(* IEC 61131-3 sources: kns-port-domestic/targets/astra/src/POUs/Station/FB_PumpRotation, 14 files *)

(* ---- FB_PumpRotation.decl.st ---- *)
// Назначение: роли насосов, чередование и ограничение непрерывной работы (04 §5, §8). Запросы
//             получают насосы с ролями Lead и Assist; роли работающих по запросу насосов
//             сохраняются; недостающая роль — сначала ReadyToStart, затем доступные в паузе,
//             внутри группы — по eRotation (RunHours, Cyclic, Fixed); в ПИД ведущим — насос со
//             связью с ПЧ. Новый запрос — не раньше tStagger после предыдущего (если тот ещё
//             запрошен). Снятие роли: RunHours — насос с большей наработкой, Cyclic/Fixed —
//             подпорный. Отказавший насос теряет запрос сразу. Передача роли с перекрытием
//             tOverlap после tMaxContRun (событие 101007), повтор через STN_HANDOVER_RETRY.
//             uiRequestLimit (последовательный пуск) ограничивает новые запросы: насосы, уже
//             работающие по запросу (подхват при старте ПЛК), им не снимаются.
// Автор:      kr0nsch
// Версия:     0.1.0
// Документ:   docs/DESIGN.md, раздел 6.5; docs/04_algorithms.md, разделы 5, 8
FUNCTION_BLOCK FB_PumpRotation
VAR_INPUT
    xEnable          : BOOL;        // станция в «Автомате» (иначе запросов нет, роли считаются)
    uiRequired       : UINT;        // от действующего управления, 0…STN_PUMP_COUNT
    uiRequestLimit   : UINT;        // FB_PowerRestore: сколько запросов можно выдать
    xRequireComm     : BOOL;        // eControlAct = LevelPid: ведущий — только со связью
    xHandoverAllowed : BOOL;        // не Emergency, Float, Restart
    xAdopt           : BOOL;        // импульс: роли получают работающие насосы (вход в «Автомат», смена управления)
    axAdoptRun       : ARRAY[1..GVL_Const.STN_PUMP_COUNT] OF BOOL;  // «работает» для xAdopt (старт: GVL_IO.xP10n_RFB)
    aitfPump         : ARRAY[1..GVL_Const.STN_PUMP_COUNT] OF PL.I_MotorVfd;
    axCommOk         : ARRAY[1..GVL_Const.STN_PUMP_COUNT] OF BOOL;
    itfTime          : PL.I_TimeSource;
    itfEvents        : I_StationEventSink;
END_VAR
VAR_IN_OUT CONSTANT
    stCfg : ST_StationCfg;          // eRotation, uiDutyMax, tMaxContRun, tOverlap, tStagger
END_VAR
VAR_IN_OUT
    stRetain : ST_StationRetain;    // uiNextLead (Cyclic)
END_VAR
VAR_OUTPUT
    axRun              : ARRAY[1..GVL_Const.STN_PUMP_COUNT] OF BOOL;   // → fbP10n.xAutoRun
    aeRole             : ARRAY[1..GVL_Const.STN_PUMP_COUNT] OF E_PumpRole;
    uiLead             : UINT;
    uiAvailable        : UINT;      // Available
    uiRunning          : UINT;      // Running в любом режиме
    uiForeign          : UINT;      // работают не в Auto (сторонние, 04 §5.1)
    uiRequests         : UINT;      // запросы: не больше MAX(0, uiRequired - uiForeign), новые — до uiRequestLimit
    uiRunningRequested : UINT;      // запрошены и работают по ОС (для FB_PowerRestore)
    xHandover          : BOOL;      // идёт передача роли (перекрытие)
    xStaggerWait       : BOOL;      // новый запрос ждёт tStagger
END_VAR
VAR
    // снимок насосов этого вызова (методы читают его, а не интерфейсы)
    axAvail       : ARRAY[1..GVL_Const.STN_PUMP_COUNT] OF BOOL;    // Available
    axRunning     : ARRAY[1..GVL_Const.STN_PUMP_COUNT] OF BOOL;    // Running
    axReady       : ARRAY[1..GVL_Const.STN_PUMP_COUNT] OF BOOL;    // ReadyToStart
    audiHours     : ARRAY[1..GVL_Const.STN_PUMP_COUNT] OF UDINT;   // RunSeconds
    audiStarts    : ARRAY[1..GVL_Const.STN_PUMP_COUNT] OF UDINT;   // Starts
    audiCurRun    : ARRAY[1..GVL_Const.STN_PUMP_COUNT] OF UDINT;   // CurrentRunSeconds
    axForeign     : ARRAY[1..GVL_Const.STN_PUMP_COUNT] OF BOOL;    // работает не в Auto
    // запросы и роли
    axReq         : ARRAY[1..GVL_Const.STN_PUMP_COUNT] OF BOOL;    // запрос (роль Lead или Assist)
    audiReqSeq    : ARRAY[1..GVL_Const.STN_PUMP_COUNT] OF UDINT;   // порядок выдачи запросов (подпорный — последний)
    udiReqSeq     : UDINT;          // счётчик выданных запросов
    uiLeadIdx     : UINT;           // ведущий; 0 — нет
    uiLeadPrev    : UINT;           // ведущий прошлого вызова (событие 101005)
    // интервал пусков
    xStaggerArmed : BOOL;           // после нового запроса идёт отсчёт tStagger
    ltLastNewReq  : LTIME;          // время последнего нового запроса
    uiLastNewPump : UINT;           // насос последнего нового запроса
    // передача роли по ограничению непрерывной работы
    xHoActive     : BOOL;           // идёт передача
    uiHoOld       : UINT;           // насос, отработавший tMaxContRun
    uiHoNew       : UINT;           // насос-замена
    uiHoTarget    : UINT;           // требуемое число насосов в момент начала передачи
    xHoRetryWait  : BOOL;           // ожидание повтора STN_HANDOVER_RETRY
    fbHoStart     : PL.FB_Delay;    // замена не пустилась за STN_HANDOVER_START_TIMEOUT
    fbHoOverlap   : PL.FB_Delay;    // перекрытие tOverlap после пуска замены
    fbHoRetry     : PL.FB_Delay;    // повтор попытки через STN_HANDOVER_RETRY
    fbSysTime     : PL.FB_SystemTime;   // запасной источник времени (itfTime = 0)
END_VAR
VAR_TEMP
    uiPump        : UINT;           // номер насоса
    uiStep        : UINT;           // шаг цикла добавления и снятия запросов
    uiPick        : UINT;           // выбранный насос
    uiCount       : UINT;           // выданных запросов
    uiTarget      : UINT;           // нужно запросов: MAX(0, uiRequired - uiForeign)
    ltNow         : LTIME;          // время этого вызова
    ePumpMode     : PL.E_DeviceMode;    // режим насоса
    xStaggerOk    : BOOL;           // новый запрос разрешён по интервалу пусков
    xHoNewRunning : BOOL;           // замена работает по ОС
    udiMaxRun_s   : UDINT;          // tMaxContRun в секундах
END_VAR

(* ---- Better.method.decl.st ---- *)
// Насос uiA предпочтительнее uiB по режиму чередования (04 §8.1); uiB = 0 — любой лучше.
// RunHours: меньше RunSeconds, затем меньше Starts, затем меньший номер; Cyclic: ближе по кругу
// к uiNext; Fixed и значение вне перечисления: меньший номер
METHOD PRIVATE Better : BOOL
VAR_INPUT
    uiA    : UINT;                  // кандидат
    uiB    : UINT;                  // лучший до него; 0 — нет
    eRot   : E_RotationMode;        // режим чередования
    uiNext : UINT;                  // Cyclic: следующий ведущий 1…STN_PUMP_COUNT
END_VAR
VAR
    uiDistA : UINT;                 // Cyclic: шагов по кругу от uiNext до uiA
    uiDistB : UINT;                 // то же до uiB
END_VAR

(* ---- Better.method.impl.st ---- *)
IF uiB = 0 THEN
    Better := TRUE;
ELSIF eRot = E_RotationMode.RunHours THEN
    IF audiHours[uiA] <> audiHours[uiB] THEN
        Better := audiHours[uiA] < audiHours[uiB];
    ELSIF audiStarts[uiA] <> audiStarts[uiB] THEN
        Better := audiStarts[uiA] < audiStarts[uiB];
    ELSE
        Better := uiA < uiB;
    END_IF
ELSIF eRot = E_RotationMode.Cyclic THEN
    uiDistA := (uiA + GVL_Const.STN_PUMP_COUNT - uiNext) MOD GVL_Const.STN_PUMP_COUNT;
    uiDistB := (uiB + GVL_Const.STN_PUMP_COUNT - uiNext) MOD GVL_Const.STN_PUMP_COUNT;
    Better := uiDistA < uiDistB;
ELSE
    Better := uiA < uiB;
END_IF

(* ---- FB_PumpRotation.impl.st ---- *)
// 0. Время вызова и снимок насосов (04 §5.1): доступные, работающие, сторонние (работают не в Auto)
IF itfTime <> 0 THEN
    ltNow := itfTime.Now();
ELSE
    ltNow := fbSysTime.Now();
END_IF
uiAvailable := 0;
uiRunning := 0;
uiForeign := 0;
FOR uiPump := 1 TO GVL_Const.STN_PUMP_COUNT DO
    IF aitfPump[uiPump] <> 0 THEN
        axAvail[uiPump] := aitfPump[uiPump].Available;
        axRunning[uiPump] := aitfPump[uiPump].Running;
        axReady[uiPump] := aitfPump[uiPump].ReadyToStart;
        audiHours[uiPump] := aitfPump[uiPump].RunSeconds;
        audiStarts[uiPump] := aitfPump[uiPump].Starts;
        audiCurRun[uiPump] := aitfPump[uiPump].CurrentRunSeconds;
        ePumpMode := aitfPump[uiPump].Mode;
    ELSE
        axAvail[uiPump] := FALSE;
        axRunning[uiPump] := FALSE;
        axReady[uiPump] := FALSE;
        audiHours[uiPump] := 0;
        audiStarts[uiPump] := 0;
        audiCurRun[uiPump] := 0;
        ePumpMode := PL.E_DeviceMode.OutOfService;
    END_IF
    IF axAvail[uiPump] THEN
        uiAvailable := uiAvailable + 1;
    END_IF
    IF axRunning[uiPump] THEN
        uiRunning := uiRunning + 1;
    END_IF
    axForeign[uiPump] := axRunning[uiPump] AND ePumpMode <> PL.E_DeviceMode.Auto;
END_FOR

// Следующий ведущий (Cyclic) вне 1…STN_PUMP_COUNT — мусор persistent-памяти: с первого насоса
IF stRetain.uiNextLead < 1 OR stRetain.uiNextLead > GVL_Const.STN_PUMP_COUNT THEN
    stRetain.uiNextLead := 1;
END_IF

udiMaxRun_s := TIME_TO_UDINT(stCfg.tMaxContRun) / GVL_Const.STN_MS_PER_S;

IF NOT xEnable THEN
    // 1. «Ручной»: запросов нет, передача роли прервана; роли считаются (Standby/None)
    FOR uiPump := 1 TO GVL_Const.STN_PUMP_COUNT DO
        axReq[uiPump] := FALSE;
    END_FOR
    uiLeadIdx := 0;
    xHoActive := FALSE;
    xHoRetryWait := FALSE;
    xStaggerArmed := FALSE;
    uiForeign := 0;
    FOR uiPump := 1 TO GVL_Const.STN_PUMP_COUNT DO
        IF axForeign[uiPump] THEN
            uiForeign := uiForeign + 1;
        END_IF
    END_FOR
    uiTarget := 0;
ELSE
    // 2. Подхват работающих насосов (вход в «Автомат», смена управления, старт ПЛК): запрос
    //    получают работающие, прежние запросы сохраняются — пуск, который ещё идёт, не обрывается.
    //    В этом вызове доступность не проверяется: устройство ещё не выполнило запрос режима
    IF xAdopt THEN
        FOR uiPump := 1 TO GVL_Const.STN_PUMP_COUNT DO
            IF axAdoptRun[uiPump] AND NOT axReq[uiPump] THEN
                axReq[uiPump] := TRUE;
                udiReqSeq := udiReqSeq + 1;
                audiReqSeq[uiPump] := udiReqSeq;
            END_IF
        END_FOR
    ELSE
        // Насос, ставший недоступным (отказ, блокировка, смена режима, нет напряжения), теряет
        // запрос сразу; после сброса он резервный (АВР — FB_Ats, 04 §9)
        FOR uiPump := 1 TO GVL_Const.STN_PUMP_COUNT DO
            IF axReq[uiPump] AND NOT axAvail[uiPump] THEN
                axReq[uiPump] := FALSE;
            END_IF
        END_FOR
    END_IF

    // 3. Ведущий снят — роль получает работающий по запросу насос (подпорный → ведущий, 04 §5.2)
    IF uiLeadIdx >= 1 AND uiLeadIdx <= GVL_Const.STN_PUMP_COUNT THEN
        IF NOT axReq[uiLeadIdx] THEN
            uiLeadIdx := 0;
        END_IF
    ELSE
        uiLeadIdx := 0;
    END_IF
    IF uiLeadIdx = 0 THEN
        uiLeadIdx := PickLead(xPreferComm := xRequireComm);
    END_IF

    // 4. ПИД: ведущий без связи, а у другого запрошенного насоса связь есть — смена ведущего без
    //    пуска и останова (оба получают одно задание частоты, 04 §12)
    IF xRequireComm AND uiLeadIdx <> 0 THEN
        IF NOT axCommOk[uiLeadIdx] THEN
            uiPick := PickLeadIn(xCommOnly := TRUE);
            IF uiPick <> 0 THEN
                uiLeadIdx := uiPick;
            END_IF
        END_IF
    END_IF

    uiCount := 0;
    FOR uiPump := 1 TO GVL_Const.STN_PUMP_COUNT DO
        IF axReq[uiPump] THEN
            uiCount := uiCount + 1;
        END_IF
    END_FOR
    // Запросов нужно: требуемое число минус сторонние работающие (04 §5.1), не меньше 0. Сторонний —
    // работает не в Auto и не запрошен станцией: подхваченный насос, который ещё не перешёл в Auto
    // (запрос режима выполнит устройство), сторонним не считается
    uiForeign := 0;
    FOR uiPump := 1 TO GVL_Const.STN_PUMP_COUNT DO
        IF axForeign[uiPump] AND NOT axReq[uiPump] THEN
            uiForeign := uiForeign + 1;
        END_IF
    END_FOR
    uiTarget := MIN(uiRequired, GVL_Const.STN_PUMP_COUNT);
    uiTarget := SEL(uiTarget > uiForeign, 0, uiTarget - uiForeign);

    // 5. Передача роли (04 §8.2): прервать, если условия изменились или замена отказала
    IF xHoActive THEN
        IF NOT xHandoverAllowed OR uiTarget <> uiHoTarget OR NOT axReq[uiHoOld] OR NOT axReq[uiHoNew] THEN
            xHoActive := FALSE;
            // замена потеряла запрос (отказ при пуске, АВР) — прежний насос работает, повтор позже
            xHoRetryWait := axReq[uiHoOld] AND NOT axReq[uiHoNew];
        END_IF
    END_IF
END_IF

// Выдержки передачи роли вызываются каждый цикл (FB_Delay должен видеть каждую смену входа)
xHoNewRunning := FALSE;
IF xHoActive AND uiHoNew >= 1 AND uiHoNew <= GVL_Const.STN_PUMP_COUNT THEN
    xHoNewRunning := axRunning[uiHoNew];
END_IF
fbHoStart(xIn := xHoActive AND NOT xHoNewRunning, tOnDelay := GVL_Const.STN_HANDOVER_START_TIMEOUT,
          itfTime := itfTime);
fbHoOverlap(xIn := xHoActive AND xHoNewRunning, tOnDelay := stCfg.tOverlap, itfTime := itfTime);

IF xEnable THEN
    IF xHoActive THEN
        IF fbHoStart.xOut THEN
            // замена не вышла в работу: запрос с неё снимается, прежний насос работает дальше
            axReq[uiHoNew] := FALSE;
            uiCount := uiCount - 1;
            xHoActive := FALSE;
            xHoRetryWait := TRUE;
        ELSIF fbHoOverlap.xOut THEN
            // замена в работе дольше tOverlap: она получает роль прежнего насоса, тот останавливается
            IF uiLeadIdx = uiHoOld THEN
                uiLeadIdx := uiHoNew;
            END_IF
            axReq[uiHoOld] := FALSE;
            uiCount := uiCount - 1;
            xHoActive := FALSE;
            IF itfEvents <> 0 THEN
                itfEvents.LogEvent(eEvent := E_StationEvent.ContRunHandover, rValue := UINT_TO_REAL(uiHoNew));
            END_IF
        END_IF
    ELSIF xHandoverAllowed AND stCfg.tMaxContRun > T#0S AND NOT xHoRetryWait AND uiCount = uiTarget THEN
        // насос с запросом работает непрерывно дольше tMaxContRun (берётся самый долгий)
        uiPick := 0;
        FOR uiPump := 1 TO GVL_Const.STN_PUMP_COUNT DO
            IF axReq[uiPump] AND axRunning[uiPump] AND audiCurRun[uiPump] >= udiMaxRun_s THEN
                IF uiPick = 0 THEN
                    uiPick := uiPump;
                ELSIF audiCurRun[uiPump] > audiCurRun[uiPick] THEN
                    uiPick := uiPump;
                END_IF
            END_IF
        END_FOR
        IF uiPick <> 0 THEN
            uiHoOld := uiPick;
            // замена — только готовый к пуску резервный; ведущему в ПИД — со связью
            uiHoNew := PickCandidate(eRot := stCfg.eRotation, uiNext := stRetain.uiNextLead,
                                     xNeedComm := xRequireComm AND uiPick = uiLeadIdx, xReadyOnly := TRUE);
            IF uiHoNew <> 0 THEN
                axReq[uiHoNew] := TRUE;
                udiReqSeq := udiReqSeq + 1;
                audiReqSeq[uiHoNew] := udiReqSeq;
                uiCount := uiCount + 1;
                xHoActive := TRUE;
                uiHoTarget := uiTarget;
                xStaggerArmed := TRUE;
                ltLastNewReq := ltNow;
                uiLastNewPump := uiHoNew;
            ELSE
                xHoRetryWait := TRUE;                       // резерва нет — повтор через STN_HANDOVER_RETRY
            END_IF
        END_IF
    END_IF

    // 6. Снятие лишних запросов (04 §5.2): RunHours — насос с большей наработкой, Cyclic/Fixed —
    //    подпорный; во время передачи роли запрос замены не лишний
    IF NOT xHoActive THEN
        FOR uiStep := 1 TO GVL_Const.STN_PUMP_COUNT DO
            IF uiCount > uiTarget THEN
                uiPick := PickToRemove(eRot := stCfg.eRotation);
                IF uiPick <> 0 THEN
                    axReq[uiPick] := FALSE;
                    uiCount := uiCount - 1;
                    IF uiPick = uiLeadIdx THEN
                        uiLeadIdx := PickLead(xPreferComm := xRequireComm);
                    END_IF
                END_IF
            END_IF
        END_FOR
    END_IF

    // 7. Новые запросы: не больше нужного, новые — не больше uiRequestLimit (последовательный пуск),
    //    по одному с интервалом tStagger, если насос предыдущего нового запроса ещё запрошен.
    //    «Время назад» — интервал отсчитывается заново (два пуска подряд не допускаются)
    IF ltNow < ltLastNewReq THEN
        ltLastNewReq := ltNow;
    END_IF
    FOR uiStep := 1 TO GVL_Const.STN_PUMP_COUNT DO
        xStaggerOk := TRUE;
        IF xStaggerArmed AND uiLastNewPump >= 1 AND uiLastNewPump <= GVL_Const.STN_PUMP_COUNT THEN
            IF axReq[uiLastNewPump] THEN
                // PORT: [types] проверить в Astra.IDE — литералы и преобразования LTIME (C11)
                xStaggerOk := ltNow - ltLastNewReq >= TIME_TO_LTIME(stCfg.tStagger);
            END_IF
        END_IF
        IF NOT xHoActive AND uiCount < uiTarget AND uiCount < uiRequestLimit AND xStaggerOk THEN
            uiPick := PickCandidate(eRot := stCfg.eRotation, uiNext := stRetain.uiNextLead,
                                    xNeedComm := xRequireComm AND uiLeadIdx = 0, xReadyOnly := FALSE);
            IF uiPick <> 0 THEN
                axReq[uiPick] := TRUE;
                udiReqSeq := udiReqSeq + 1;
                audiReqSeq[uiPick] := udiReqSeq;
                uiCount := uiCount + 1;
                xStaggerArmed := TRUE;
                ltLastNewReq := ltNow;
                uiLastNewPump := uiPick;
                IF uiLeadIdx = 0 THEN
                    // новый ведущий; по кругу — следующий после него (энергонезависимо)
                    uiLeadIdx := uiPick;
                    IF stCfg.eRotation = E_RotationMode.Cyclic THEN
                        stRetain.uiNextLead := (uiPick MOD GVL_Const.STN_PUMP_COUNT) + 1;
                    END_IF
                END_IF
            END_IF
        END_IF
    END_FOR

    // ожидание интервала пусков (HMI): нужен ещё насос, кандидат есть, но tStagger не истёк
    xStaggerOk := TRUE;
    IF xStaggerArmed AND uiLastNewPump >= 1 AND uiLastNewPump <= GVL_Const.STN_PUMP_COUNT THEN
        IF axReq[uiLastNewPump] THEN
            // PORT: [types] проверить в Astra.IDE — литералы и преобразования LTIME (C11)
            xStaggerOk := ltNow - ltLastNewReq >= TIME_TO_LTIME(stCfg.tStagger);
        END_IF
    END_IF
    xStaggerWait := FALSE;
    IF NOT xHoActive AND uiCount < uiTarget AND uiCount < uiRequestLimit AND NOT xStaggerOk THEN
        xStaggerWait := PickCandidate(eRot := stCfg.eRotation, uiNext := stRetain.uiNextLead,
                                      xNeedComm := FALSE, xReadyOnly := FALSE) <> 0;
    END_IF
ELSE
    xStaggerWait := FALSE;
END_IF

fbHoRetry(xIn := xHoRetryWait, tOnDelay := GVL_Const.STN_HANDOVER_RETRY, itfTime := itfTime);
IF fbHoRetry.xOut THEN
    xHoRetryWait := FALSE;
END_IF

// 8. Выходы: запросы, роли (04 §5.1), счётчики; событие смены ведущего (101005, номер насоса)
uiRequests := 0;
uiRunningRequested := 0;
FOR uiPump := 1 TO GVL_Const.STN_PUMP_COUNT DO
    axRun[uiPump] := axReq[uiPump];
    IF axReq[uiPump] THEN
        uiRequests := uiRequests + 1;
        IF axRunning[uiPump] THEN
            uiRunningRequested := uiRunningRequested + 1;
        END_IF
        IF uiPump = uiLeadIdx THEN
            aeRole[uiPump] := E_PumpRole.Lead;
        ELSE
            aeRole[uiPump] := E_PumpRole.Assist;
        END_IF
    ELSIF axAvail[uiPump] THEN
        aeRole[uiPump] := E_PumpRole.Standby;
    ELSE
        aeRole[uiPump] := E_PumpRole.None;
    END_IF
END_FOR
uiLead := uiLeadIdx;
xHandover := xHoActive;
// По кругу следующий ведущий отсчитывается от любого нового ведущего — и без пуска (передача роли, подпорный
// стал ведущим, подхват): иначе тот же насос снова получил бы следующий пуск (04 §8.1)
IF uiLeadIdx <> uiLeadPrev AND uiLeadIdx <> 0 THEN
    IF stCfg.eRotation = E_RotationMode.Cyclic THEN
        stRetain.uiNextLead := (uiLeadIdx MOD GVL_Const.STN_PUMP_COUNT) + 1;
    END_IF
    IF itfEvents <> 0 THEN
        itfEvents.LogEvent(eEvent := E_StationEvent.LeadChanged, rValue := UINT_TO_REAL(uiLeadIdx));
    END_IF
END_IF
uiLeadPrev := uiLeadIdx;

(* ---- PickCandidate.method.decl.st ---- *)
// Насос для нового запроса (04 §5.2): сначала ReadyToStart, затем доступные в паузе (tMinStop,
// лимит пусков: запрос подождёт); внутри группы — по режиму чередования. xNeedComm — назначается
// ведущий в ПИД: сначала насосы со связью с ПЧ; если таких нет, — любой (станция откачивает, ПИД
// без связи не готов, и действует ступенчатое, 04 §12); при передаче роли (xReadyOnly) — только со связью.
// 0 — кандидата нет
METHOD PRIVATE PickCandidate : UINT
VAR_INPUT
    eRot       : E_RotationMode;        // режим чередования
    uiNext     : UINT;                  // Cyclic: следующий ведущий
    xNeedComm  : BOOL;                  // предпочесть насосы со связью
    xReadyOnly : BOOL;                  // только готовые к пуску (передача роли)
END_VAR

(* ---- PickCandidate.method.impl.st ---- *)
PickCandidate := 0;
IF xNeedComm THEN
    PickCandidate := PickIn(eRot := eRot, uiNext := uiNext, xRequireCommOk := TRUE, xRequireReady := TRUE);
    IF PickCandidate = 0 AND NOT xReadyOnly THEN
        PickCandidate := PickIn(eRot := eRot, uiNext := uiNext, xRequireCommOk := TRUE, xRequireReady := FALSE);
    END_IF
END_IF
// передача роли ведущего в ПИД — только насосу со связью: без неё после перекрытия ПИД потерял бы готовность
// и станция ушла бы в ступенчатое (04 §5.2 п. 3); нет такого — повтор передачи позже
IF PickCandidate = 0 AND NOT (xNeedComm AND xReadyOnly) THEN
    PickCandidate := PickIn(eRot := eRot, uiNext := uiNext, xRequireCommOk := FALSE, xRequireReady := TRUE);
    IF PickCandidate = 0 AND NOT xReadyOnly THEN
        PickCandidate := PickIn(eRot := eRot, uiNext := uiNext, xRequireCommOk := FALSE, xRequireReady := FALSE);
    END_IF
END_IF

(* ---- PickIn.method.decl.st ---- *)
// Лучший незапрошенный доступный насос группы по режиму чередования; 0 — нет такого.
// xRequireReady — только ReadyToStart, xRequireCommOk — только со связью с ПЧ
METHOD PRIVATE PickIn : UINT
VAR_INPUT
    eRot           : E_RotationMode;    // режим чередования
    uiNext         : UINT;              // Cyclic: следующий ведущий
    xRequireCommOk : BOOL;              // только насосы со связью
    xRequireReady  : BOOL;              // только готовые к пуску
END_VAR
VAR
    uiIdx : UINT;                       // номер насоса
END_VAR

(* ---- PickIn.method.impl.st ---- *)
PickIn := 0;
FOR uiIdx := 1 TO GVL_Const.STN_PUMP_COUNT DO
    IF NOT axReq[uiIdx] AND axAvail[uiIdx] AND (axReady[uiIdx] OR NOT xRequireReady)
       AND (axCommOk[uiIdx] OR NOT xRequireCommOk) THEN
        IF Better(uiA := uiIdx, uiB := PickIn, eRot := eRot, uiNext := uiNext) THEN
            PickIn := uiIdx;
        END_IF
    END_IF
END_FOR

(* ---- PickLead.method.decl.st ---- *)
// Ведущий среди запрошенных насосов; xPreferComm (ПИД) — сначала насосы со связью с ПЧ, если
// таких нет — любой запрошенный. 0 — нет запрошенных
METHOD PRIVATE PickLead : UINT
VAR_INPUT
    xPreferComm : BOOL;                 // предпочесть насосы со связью
END_VAR

(* ---- PickLead.method.impl.st ---- *)
PickLead := 0;
IF xPreferComm THEN
    PickLead := PickLeadIn(xCommOnly := TRUE);
END_IF
IF PickLead = 0 THEN
    PickLead := PickLeadIn(xCommOnly := FALSE);
END_IF

(* ---- PickLeadIn.method.decl.st ---- *)
// Ведущий среди запрошенных насосов: меньше наработка (04 §3.2: при подхвате ведущий — работающий
// с меньшей наработкой; 04 §5.2: после останова ведущего роль у оставшегося), затем меньше пусков,
// затем меньший номер. xCommOnly — только насосы со связью с ПЧ. 0 — нет запрошенных
METHOD PRIVATE PickLeadIn : UINT
VAR_INPUT
    xCommOnly : BOOL;                   // только со связью
END_VAR
VAR
    uiIdx : UINT;                       // номер насоса
END_VAR

(* ---- PickLeadIn.method.impl.st ---- *)
PickLeadIn := 0;
FOR uiIdx := 1 TO GVL_Const.STN_PUMP_COUNT DO
    IF axReq[uiIdx] AND (axCommOk[uiIdx] OR NOT xCommOnly) THEN
        IF Better(uiA := uiIdx, uiB := PickLeadIn, eRot := E_RotationMode.RunHours, uiNext := 1) THEN
            PickLeadIn := uiIdx;
        END_IF
    END_IF
END_FOR

(* ---- PickToRemove.method.decl.st ---- *)
// Насос, с которого снимается запрос, когда нужно меньше насосов (04 §5.2): RunHours — с большей
// наработкой (затем больше пусков, затем больший номер), Cyclic и Fixed — подпорный, выданный
// последним; ведущий — только если подпорных нет. В ПИД (xRequireComm) насос со связью с ПЧ снимается
// последним: остаться должен насос, которым ПИД может управлять (04 §5.2 п. 3). 0 — нет запрошенных
METHOD PRIVATE PickToRemove : UINT
VAR_INPUT
    eRot : E_RotationMode;              // режим чередования
END_VAR
VAR
    uiIdx      : UINT;                  // номер насоса
    uiPass     : UINT;                  // проход: 1 — только насосы без связи (ПИД), 2 — все
    xCommFirst : BOOL;                  // ПИД и есть запрошенный насос без связи
END_VAR

(* ---- PickToRemove.method.impl.st ---- *)
PickToRemove := 0;
xCommFirst := FALSE;
IF xRequireComm THEN
    FOR uiIdx := 1 TO GVL_Const.STN_PUMP_COUNT DO
        xCommFirst := xCommFirst OR (axReq[uiIdx] AND NOT axCommOk[uiIdx]);
    END_FOR
END_IF
FOR uiPass := SEL(xCommFirst, 2, 1) TO 2 DO
    IF PickToRemove = 0 THEN
        FOR uiIdx := 1 TO GVL_Const.STN_PUMP_COUNT DO
            IF axReq[uiIdx] AND (uiPass = 2 OR NOT axCommOk[uiIdx]) THEN
                IF eRot = E_RotationMode.RunHours THEN
                    // наоборот к выбору при пуске: насос, который проигрывает всем остальным
                    IF PickToRemove = 0 THEN
                        PickToRemove := uiIdx;
                    ELSIF Better(uiA := PickToRemove, uiB := uiIdx, eRot := eRot, uiNext := 1) THEN
                        PickToRemove := uiIdx;
                    END_IF
                ELSIF uiIdx <> uiLeadIdx THEN
                    IF PickToRemove = 0 THEN
                        PickToRemove := uiIdx;
                    ELSIF audiReqSeq[uiIdx] > audiReqSeq[PickToRemove] THEN
                        PickToRemove := uiIdx;
                    END_IF
                END_IF
            END_IF
        END_FOR
    END_IF
END_FOR
IF PickToRemove = 0 AND uiLeadIdx >= 1 AND uiLeadIdx <= GVL_Const.STN_PUMP_COUNT THEN
    IF axReq[uiLeadIdx] THEN
        PickToRemove := uiLeadIdx;
    END_IF
END_IF
